// TIA Portal V18 export
FUNCTION "BYPASS DOS EQUIPAMENTOS" : Void   // FC12, LAD
{ S7_Optimized_Access := 'TRUE' }
// stored: SetENOAutomatically false
BEGIN

REGION Network 1: BYPASS GERAL E ESVAZIAMENTO DOS TRANSPORTADORES
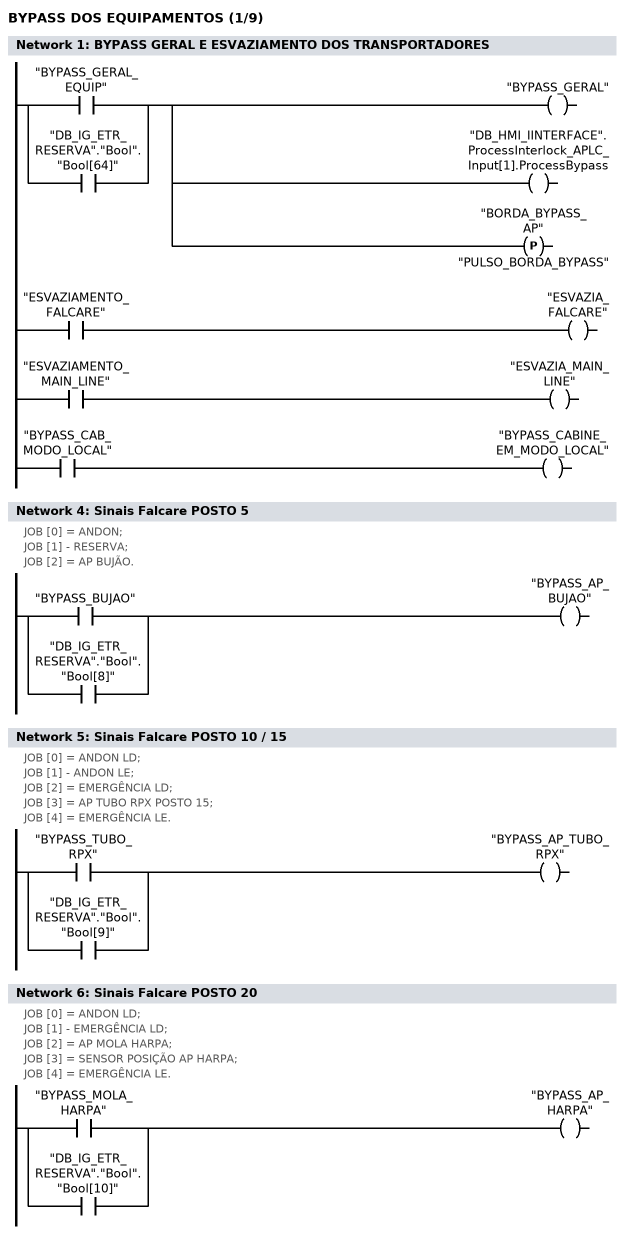
   "BYPASS_GERAL" := "BYPASS_GERAL_EQUIP" OR "DB_IG_ETR_RESERVA"."Bool"."Bool[64]";
   "DB_HMI_IINTERFACE".ProcessInterlock_APLC_Input[1].ProcessBypass := "BYPASS_GERAL";
   "BORDA_BYPASS_AP" := "BYPASS_GERAL" AND NOT "PULSO_BORDA_BYPASS";   // rising edge
   "PULSO_BORDA_BYPASS" := "BYPASS_GERAL";
   "ESVAZIA_FALCARE" := "ESVAZIAMENTO_FALCARE";
   "ESVAZIA_MAIN_LINE" := "ESVAZIAMENTO_MAIN_LINE";
   "BYPASS_CABINE_EM_MODO_LOCAL" := "BYPASS_CAB_MODO_LOCAL";
END_REGION

REGION Network 2: Sinais Falcare POSTO 1
   // JOB [0] = ANDON;
   // JOB [1] - EMERGÊNCIA;
END_REGION

REGION Network 3: Sinais Falcare VIVERK
   // JOB [0] = ANDON;
   // JOB [1] - EMERGÊNCIA;
END_REGION

REGION Network 4: Sinais Falcare POSTO 5
   // JOB [0] = ANDON;
   // JOB [1] - RESERVA;
   // JOB [2] = AP BUJÃO.
   RUNG wire#powerrail
      Contact( "BYPASS_BUJAO" )
      wire#w1
      Coil( "BYPASS_AP_BUJAO" )
   END_RUNG
   RUNG wire#powerrail
      Contact( "DB_IG_ETR_RESERVA"."Bool"."Bool[8]" )
   END_RUNG wire#w1
   // the same network as SCL:
   "BYPASS_AP_BUJAO" := "BYPASS_BUJAO" OR "DB_IG_ETR_RESERVA"."Bool"."Bool[8]";
END_REGION

REGION Network 5: Sinais Falcare POSTO 10 / 15
   // JOB [0] = ANDON LD;
   // JOB [1] - ANDON LE;
   // JOB [2] = EMERGÊNCIA LD;
   // JOB [3] = AP TUBO RPX POSTO 15;
   // JOB [4] = EMERGÊNCIA LE.
   RUNG wire#powerrail
      Contact( "BYPASS_TUBO_RPX" )
      wire#w1
      Coil( "BYPASS_AP_TUBO_RPX" )
   END_RUNG
   RUNG wire#powerrail
      Contact( "DB_IG_ETR_RESERVA"."Bool"."Bool[9]" )
   END_RUNG wire#w1
   // the same network as SCL:
   "BYPASS_AP_TUBO_RPX" := "BYPASS_TUBO_RPX" OR "DB_IG_ETR_RESERVA"."Bool"."Bool[9]";
END_REGION

REGION Network 6: Sinais Falcare POSTO 20
   // JOB [0] = ANDON LD;
   // JOB [1] - EMERGÊNCIA LD;
   // JOB [2] = AP MOLA HARPA;
   // JOB [3] = SENSOR POSIÇÃO AP HARPA;
   // JOB [4] = EMERGÊNCIA LE.
   RUNG wire#powerrail
      Contact( "BYPASS_MOLA_HARPA" )
      wire#w1
      Coil( "BYPASS_AP_HARPA" )
   END_RUNG
   RUNG wire#powerrail
      Contact( "DB_IG_ETR_RESERVA"."Bool"."Bool[10]" )
   END_RUNG wire#w1
   // the same network as SCL:
   "BYPASS_AP_HARPA" := "BYPASS_MOLA_HARPA" OR "DB_IG_ETR_RESERVA"."Bool"."Bool[10]";
END_REGION

REGION Network 7: Sinais Falcare POSTO 30
   // JOB [0] = ANDON LD;
   // JOB [1] = ANDON LE;
   // JOB [2] = EMERGENCIA;
   // JOB [3] = AP DA CARCAÇA;
   // JOB [4] = POSIÇÃO TALHA DIF.
   // JOB [5] = PY JUNTA.
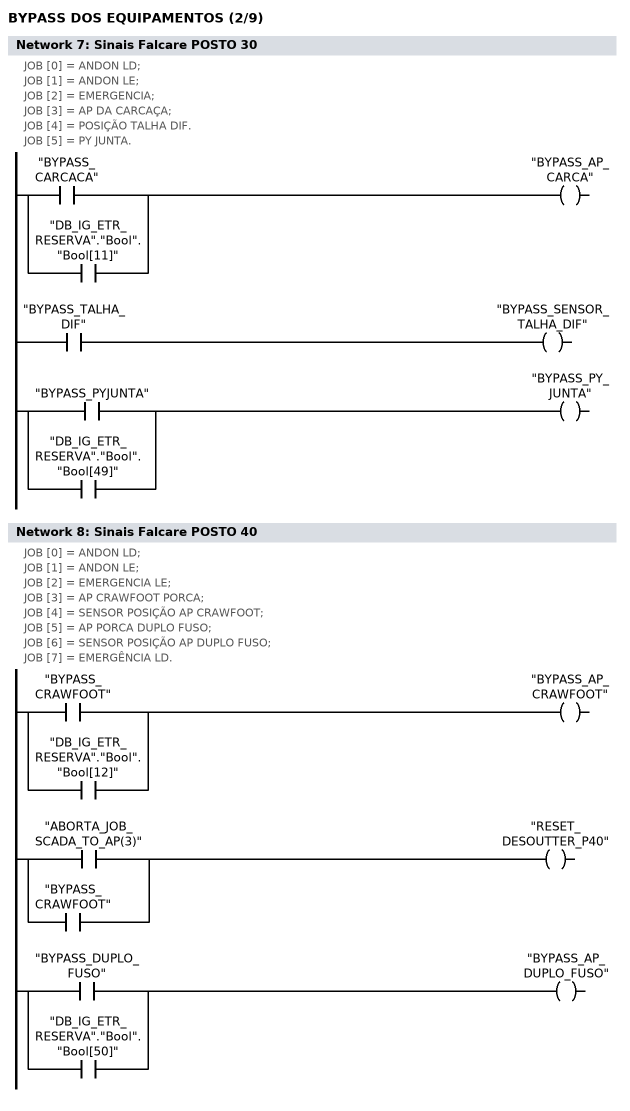
   RUNG wire#powerrail
      Contact( "BYPASS_CARCACA" )
      wire#w1
      Coil( "BYPASS_AP_CARCA" )
   END_RUNG
   RUNG wire#powerrail
      Contact( "DB_IG_ETR_RESERVA"."Bool"."Bool[11]" )
   END_RUNG wire#w1
   RUNG wire#powerrail
      Contact( "BYPASS_TALHA_DIF" )
      Coil( "BYPASS_SENSOR_TALHA_DIF" )
   END_RUNG
   RUNG wire#powerrail
      Contact( "BYPASS_PYJUNTA" )
      wire#w2
      Coil( "BYPASS_PY_JUNTA" )
   END_RUNG
   RUNG wire#powerrail
      Contact( "DB_IG_ETR_RESERVA"."Bool"."Bool[49]" )
   END_RUNG wire#w2
   // the same network as SCL:
   "BYPASS_AP_CARCA" := "BYPASS_CARCACA" OR "DB_IG_ETR_RESERVA"."Bool"."Bool[11]";
   "BYPASS_SENSOR_TALHA_DIF" := "BYPASS_TALHA_DIF";
   "BYPASS_PY_JUNTA" := "BYPASS_PYJUNTA" OR "DB_IG_ETR_RESERVA"."Bool"."Bool[49]";
END_REGION

REGION Network 8: Sinais Falcare POSTO 40
   // JOB [0] = ANDON LD;
   // JOB [1] = ANDON LE;
   // JOB [2] = EMERGENCIA LE;
   // JOB [3] = AP CRAWFOOT PORCA;
   // JOB [4] = SENSOR POSIÇÃO AP CRAWFOOT;
   // JOB [5] = AP PORCA DUPLO FUSO;
   // JOB [6] = SENSOR POSIÇÃO AP DUPLO FUSO;
   // JOB [7] = EMERGÊNCIA LD.
   RUNG wire#powerrail
      Contact( "BYPASS_CRAWFOOT" )
      wire#w1
      Coil( "BYPASS_AP_CRAWFOOT" )
   END_RUNG
   RUNG wire#powerrail
      Contact( "DB_IG_ETR_RESERVA"."Bool"."Bool[12]" )
   END_RUNG wire#w1
   RUNG wire#powerrail
      Contact( "ABORTA_JOB_SCADA_TO_AP(3)" )
      wire#w2
      Coil( "RESET_DESOUTTER_P40" )
   END_RUNG
   RUNG wire#powerrail
      Contact( "BYPASS_CRAWFOOT" )
   END_RUNG wire#w2
   RUNG wire#powerrail
      Contact( "BYPASS_DUPLO_FUSO" )
      wire#w3
      Coil( "BYPASS_AP_DUPLO_FUSO" )
   END_RUNG
   RUNG wire#powerrail
      Contact( "DB_IG_ETR_RESERVA"."Bool"."Bool[50]" )
   END_RUNG wire#w3
   // the same network as SCL:
   "BYPASS_AP_CRAWFOOT" := "BYPASS_CRAWFOOT" OR "DB_IG_ETR_RESERVA"."Bool"."Bool[12]";
   "RESET_DESOUTTER_P40" := "ABORTA_JOB_SCADA_TO_AP(3)" OR "BYPASS_CRAWFOOT";
   "BYPASS_AP_DUPLO_FUSO" := "BYPASS_DUPLO_FUSO" OR "DB_IG_ETR_RESERVA"."Bool"."Bool[50]";
END_REGION

REGION Network 9: Sinais Falcare POSTO 50 /55
   // JOB [0] = ANDON;
   // JOB [1] = EMERGENCIA;
   // JOB [2] = AP PORCA ESCONDIDA;
   // JOB [3] = SENSOR POSIÇÃO AP PORCA ESCONDIDA;
   // JOB [4] = AP PORCA SUPORTE DO CILINDRO;
   // JOB [5] = SENSOR POSIÇÃO AP SUPORTE DO CILINDRO;
   // JOB [6] = ANDON LD.
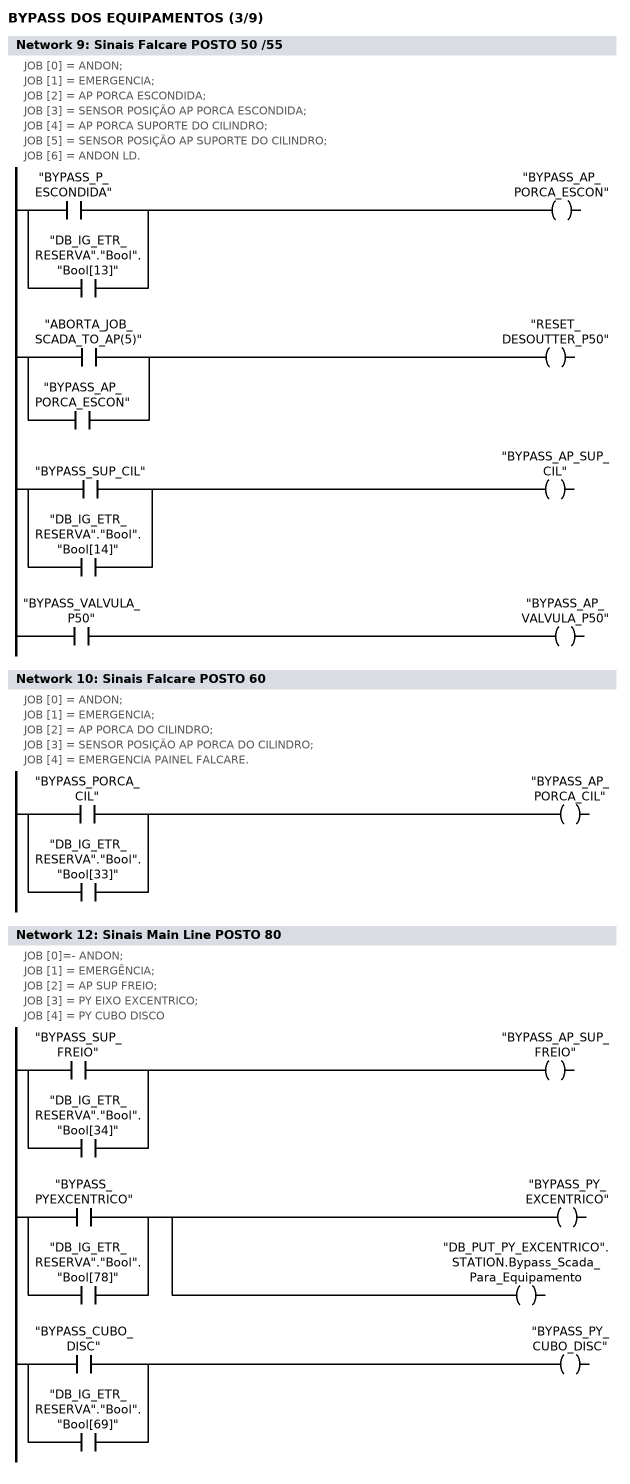
   RUNG wire#powerrail
      Contact( "BYPASS_P_ESCONDIDA" )
      wire#w1
      Coil( "BYPASS_AP_PORCA_ESCON" )
   END_RUNG
   RUNG wire#powerrail
      Contact( "DB_IG_ETR_RESERVA"."Bool"."Bool[13]" )
   END_RUNG wire#w1
   RUNG wire#powerrail
      Contact( "ABORTA_JOB_SCADA_TO_AP(5)" )
      wire#w2
      Coil( "RESET_DESOUTTER_P50" )
   END_RUNG
   RUNG wire#powerrail
      Contact( "BYPASS_AP_PORCA_ESCON" )
   END_RUNG wire#w2
   RUNG wire#powerrail
      Contact( "BYPASS_SUP_CIL" )
      wire#w3
      Coil( "BYPASS_AP_SUP_CIL" )
   END_RUNG
   RUNG wire#powerrail
      Contact( "DB_IG_ETR_RESERVA"."Bool"."Bool[14]" )
   END_RUNG wire#w3
   RUNG wire#powerrail
      Contact( "BYPASS_VALVULA_P50" )
      Coil( "BYPASS_AP_VALVULA_P50" )
   END_RUNG
   // the same network as SCL:
   "BYPASS_AP_PORCA_ESCON" := "BYPASS_P_ESCONDIDA" OR "DB_IG_ETR_RESERVA"."Bool"."Bool[13]";
   "RESET_DESOUTTER_P50" := "ABORTA_JOB_SCADA_TO_AP(5)" OR "BYPASS_AP_PORCA_ESCON";
   "BYPASS_AP_SUP_CIL" := "BYPASS_SUP_CIL" OR "DB_IG_ETR_RESERVA"."Bool"."Bool[14]";
   "BYPASS_AP_VALVULA_P50" := "BYPASS_VALVULA_P50";
END_REGION

REGION Network 10: Sinais Falcare POSTO 60
   // JOB [0] = ANDON;
   // JOB [1] = EMERGENCIA;
   // JOB [2] = AP PORCA DO CILINDRO;
   // JOB [3] = SENSOR POSIÇÃO AP PORCA DO CILINDRO;
   // JOB [4] = EMERGENCIA PAINEL FALCARE.
   RUNG wire#powerrail
      Contact( "BYPASS_PORCA_CIL" )
      wire#w1
      Coil( "BYPASS_AP_PORCA_CIL" )
   END_RUNG
   RUNG wire#powerrail
      Contact( "DB_IG_ETR_RESERVA"."Bool"."Bool[33]" )
   END_RUNG wire#w1
   // the same network as SCL:
   "BYPASS_AP_PORCA_CIL" := "BYPASS_PORCA_CIL" OR "DB_IG_ETR_RESERVA"."Bool"."Bool[33]";
END_REGION

REGION Network 11: Sinais Main Line POSTO 70 / 75
   // \\ JOB [0] - ANDON
END_REGION

REGION Network 12: Sinais Main Line POSTO 80
   // JOB [0]=- ANDON;
   // JOB [1] = EMERGÊNCIA;
   // JOB [2] = AP SUP FREIO;
   // JOB [3] = PY EIXO EXCENTRICO;
   // JOB [4] = PY CUBO DISCO
   RUNG wire#powerrail
      Contact( "BYPASS_SUP_FREIO" )
      wire#w1
      Coil( "BYPASS_AP_SUP_FREIO" )
   END_RUNG
   RUNG wire#powerrail
      Contact( "DB_IG_ETR_RESERVA"."Bool"."Bool[34]" )
   END_RUNG wire#w1
   RUNG wire#powerrail
      Contact( "BYPASS_PYEXCENTRICO" )
      wire#w2
      Coil( "BYPASS_PY_EXCENTRICO" )
   END_RUNG
   RUNG wire#powerrail
      Contact( "DB_IG_ETR_RESERVA"."Bool"."Bool[78]" )
   END_RUNG wire#w2
   RUNG wire#w2
      Coil( "DB_PUT_PY_EXCENTRICO".STATION.Bypass_Scada_Para_Equipamento )
   END_RUNG
   RUNG wire#powerrail
      Contact( "BYPASS_CUBO_DISC" )
      wire#w3
      Coil( "BYPASS_PY_CUBO_DISC" )
   END_RUNG
   RUNG wire#powerrail
      Contact( "DB_IG_ETR_RESERVA"."Bool"."Bool[69]" )
   END_RUNG wire#w3
   // the same network as SCL:
   "BYPASS_AP_SUP_FREIO" := "BYPASS_SUP_FREIO" OR "DB_IG_ETR_RESERVA"."Bool"."Bool[34]";
   "BYPASS_PY_EXCENTRICO" := "BYPASS_PYEXCENTRICO" OR "DB_IG_ETR_RESERVA"."Bool"."Bool[78]";
   "DB_PUT_PY_EXCENTRICO".STATION.Bypass_Scada_Para_Equipamento := "BYPASS_PY_EXCENTRICO";
   "BYPASS_PY_CUBO_DISC" := "BYPASS_CUBO_DISC" OR "DB_IG_ETR_RESERVA"."Bool"."Bool[69]";
END_REGION

REGION Network 13: Sinais Main Line POSTO 90 / 95
   // JOB [0] = ANDON;
   // JOB [1] = EMERGÊNCIA;
   // JOB [2] = AP HOLDER.
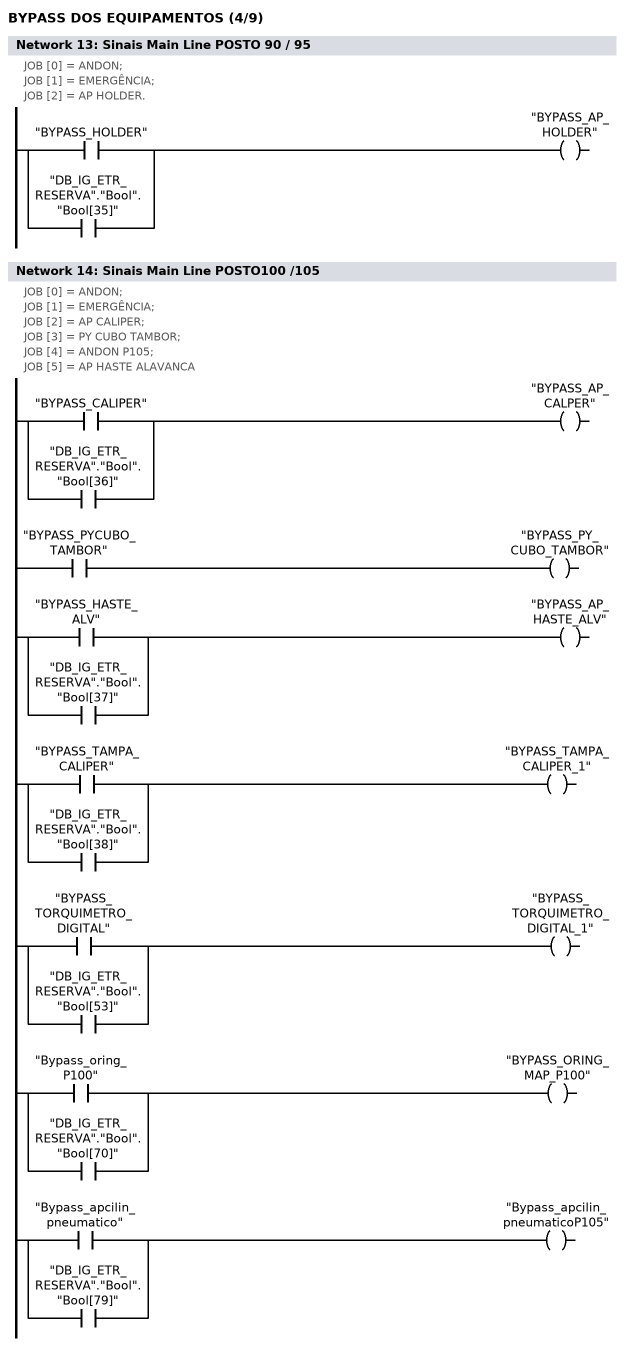
   RUNG wire#powerrail
      Contact( "BYPASS_HOLDER" )
      wire#w1
      Coil( "BYPASS_AP_HOLDER" )
   END_RUNG
   RUNG wire#powerrail
      Contact( "DB_IG_ETR_RESERVA"."Bool"."Bool[35]" )
   END_RUNG wire#w1
   // the same network as SCL:
   "BYPASS_AP_HOLDER" := "BYPASS_HOLDER" OR "DB_IG_ETR_RESERVA"."Bool"."Bool[35]";
END_REGION

REGION Network 14: Sinais Main Line POSTO100 /105
   // JOB [0] = ANDON;
   // JOB [1] = EMERGÊNCIA;
   // JOB [2] = AP CALIPER;
   // JOB [3] = PY CUBO TAMBOR;
   // JOB [4] = ANDON P105;
   // JOB [5] = AP HASTE ALAVANCA
   RUNG wire#powerrail
      Contact( "BYPASS_CALIPER" )
      wire#w1
      Coil( "BYPASS_AP_CALPER" )
   END_RUNG
   RUNG wire#powerrail
      Contact( "DB_IG_ETR_RESERVA"."Bool"."Bool[36]" )
   END_RUNG wire#w1
   RUNG wire#powerrail
      Contact( "BYPASS_PYCUBO_TAMBOR" )
      Coil( "BYPASS_PY_CUBO_TAMBOR" )
   END_RUNG
   RUNG wire#powerrail
      Contact( "BYPASS_HASTE_ALV" )
      wire#w2
      Coil( "BYPASS_AP_HASTE_ALV" )
   END_RUNG
   RUNG wire#powerrail
      Contact( "DB_IG_ETR_RESERVA"."Bool"."Bool[37]" )
   END_RUNG wire#w2
   RUNG wire#powerrail
      Contact( "BYPASS_TAMPA_CALIPER" )
      wire#w3
      Coil( "BYPASS_TAMPA_CALIPER_1" )
   END_RUNG
   RUNG wire#powerrail
      Contact( "DB_IG_ETR_RESERVA"."Bool"."Bool[38]" )
   END_RUNG wire#w3
   RUNG wire#powerrail
      Contact( "BYPASS_TORQUIMETRO_DIGITAL" )
      wire#w4
      Coil( "BYPASS_TORQUIMETRO_DIGITAL_1" )
   END_RUNG
   RUNG wire#powerrail
      Contact( "DB_IG_ETR_RESERVA"."Bool"."Bool[53]" )
   END_RUNG wire#w4
   RUNG wire#powerrail
      Contact( "Bypass_oring_P100" )
      wire#w5
      Coil( "BYPASS_ORING_MAP_P100" )
   END_RUNG
   RUNG wire#powerrail
      Contact( "DB_IG_ETR_RESERVA"."Bool"."Bool[70]" )
   END_RUNG wire#w5
   RUNG wire#powerrail
      Contact( "Bypass_apcilin_pneumatico" )
      wire#w6
      Coil( "Bypass_apcilin_pneumaticoP105" )
   END_RUNG
   RUNG wire#powerrail
      Contact( "DB_IG_ETR_RESERVA"."Bool"."Bool[79]" )
   END_RUNG wire#w6
   // the same network as SCL:
   "BYPASS_AP_CALPER" := "BYPASS_CALIPER" OR "DB_IG_ETR_RESERVA"."Bool"."Bool[36]";
   "BYPASS_PY_CUBO_TAMBOR" := "BYPASS_PYCUBO_TAMBOR";
   "BYPASS_AP_HASTE_ALV" := "BYPASS_HASTE_ALV" OR "DB_IG_ETR_RESERVA"."Bool"."Bool[37]";
   "BYPASS_TAMPA_CALIPER_1" := "BYPASS_TAMPA_CALIPER" OR "DB_IG_ETR_RESERVA"."Bool"."Bool[38]";
   "BYPASS_TORQUIMETRO_DIGITAL_1" := "BYPASS_TORQUIMETRO_DIGITAL" OR "DB_IG_ETR_RESERVA"."Bool"."Bool[53]";
   "BYPASS_ORING_MAP_P100" := "Bypass_oring_P100" OR "DB_IG_ETR_RESERVA"."Bool"."Bool[70]";
   "Bypass_apcilin_pneumaticoP105" := "Bypass_apcilin_pneumatico" OR "DB_IG_ETR_RESERVA"."Bool"."Bool[79]";
END_REGION

REGION Network 15: Sinais Main Line POSTO110 /115
   // JOB [0] = ANDON;
   // JOB [1] = SEG. BLOQUEIO CLP;
   // JOB [2] = AP CUBO;
   // JOB [3] = ANDON P115;
   // JOB [4] = CRAVADOR.
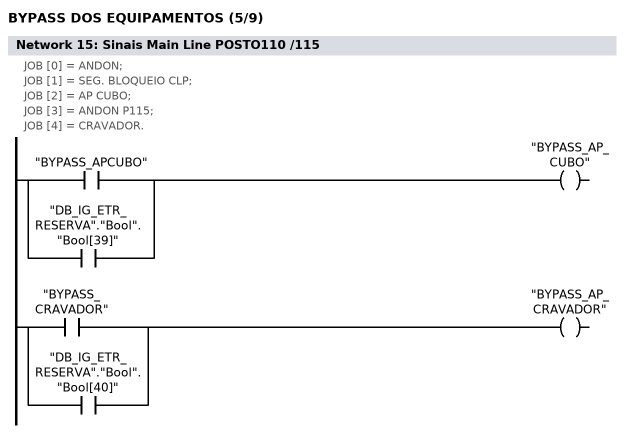
   RUNG wire#powerrail
      Contact( "BYPASS_APCUBO" )
      wire#w1
      Coil( "BYPASS_AP_CUBO" )
   END_RUNG
   RUNG wire#powerrail
      Contact( "DB_IG_ETR_RESERVA"."Bool"."Bool[39]" )
   END_RUNG wire#w1
   RUNG wire#powerrail
      Contact( "BYPASS_CRAVADOR" )
      wire#w2
      Coil( "BYPASS_AP_CRAVADOR" )
   END_RUNG
   RUNG wire#powerrail
      Contact( "DB_IG_ETR_RESERVA"."Bool"."Bool[40]" )
   END_RUNG wire#w2
   // the same network as SCL:
   "BYPASS_AP_CUBO" := "BYPASS_APCUBO" OR "DB_IG_ETR_RESERVA"."Bool"."Bool[39]";
   "BYPASS_AP_CRAVADOR" := "BYPASS_CRAVADOR" OR "DB_IG_ETR_RESERVA"."Bool"."Bool[40]";
END_REGION

REGION Network 16: Sinais Main Line POSTO120 /125
   // JOB [0] = ANDON;
   // JOB [1] - EMERGÊNCIA;
   // JOB [2] = AP INDICADOR;
   // JOB [3] = AP VALVULA;
   // JOB [4] = PY HELGE;
   // JOB [5] - ANDON P125;
   // JOB [6] - AP PORCA TERMINAL;
   // JOB [7] - AP FILTRO OLEO.
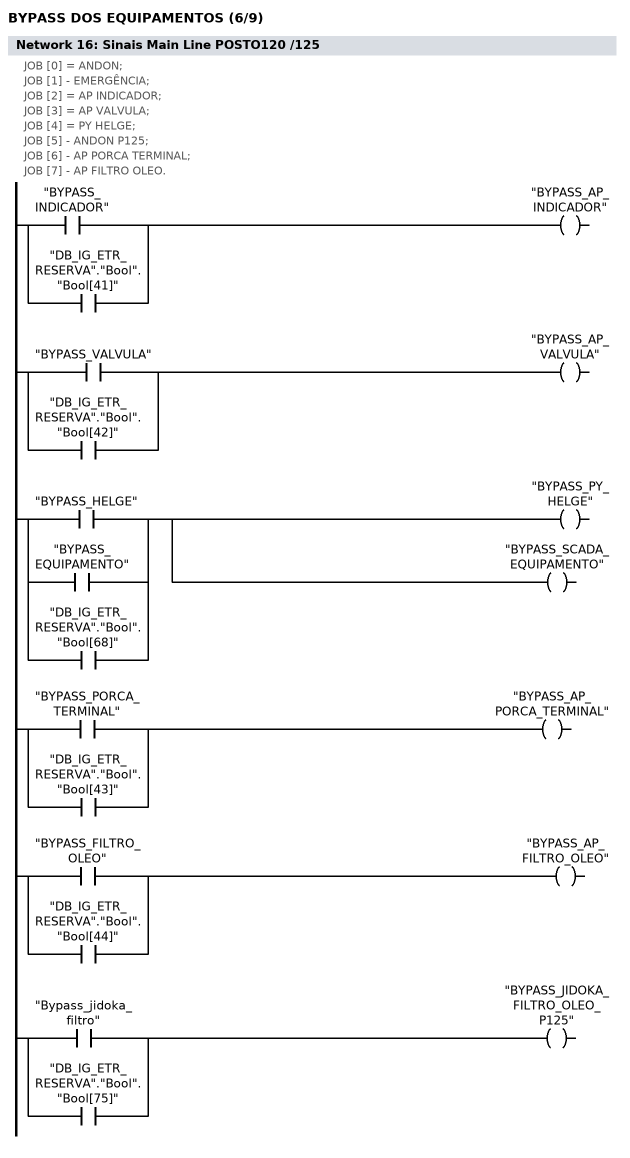
   RUNG wire#powerrail
      Contact( "BYPASS_INDICADOR" )
      wire#w1
      Coil( "BYPASS_AP_INDICADOR" )
   END_RUNG
   RUNG wire#powerrail
      Contact( "DB_IG_ETR_RESERVA"."Bool"."Bool[41]" )
   END_RUNG wire#w1
   RUNG wire#powerrail
      Contact( "BYPASS_VALVULA" )
      wire#w2
      Coil( "BYPASS_AP_VALVULA" )
   END_RUNG
   RUNG wire#powerrail
      Contact( "DB_IG_ETR_RESERVA"."Bool"."Bool[42]" )
   END_RUNG wire#w2
   RUNG wire#powerrail
      Contact( "BYPASS_HELGE" )
      wire#w3
      Coil( "BYPASS_PY_HELGE" )
   END_RUNG
   RUNG wire#powerrail
      Contact( "BYPASS_EQUIPAMENTO" )
   END_RUNG wire#w3
   RUNG wire#powerrail
      Contact( "DB_IG_ETR_RESERVA"."Bool"."Bool[68]" )
   END_RUNG wire#w3
   RUNG wire#w3
      Coil( "BYPASS_SCADA_EQUIPAMENTO" )
   END_RUNG
   RUNG wire#powerrail
      Contact( "BYPASS_PORCA_TERMINAL" )
      wire#w4
      Coil( "BYPASS_AP_PORCA_TERMINAL" )
   END_RUNG
   RUNG wire#powerrail
      Contact( "DB_IG_ETR_RESERVA"."Bool"."Bool[43]" )
   END_RUNG wire#w4
   RUNG wire#powerrail
      Contact( "BYPASS_FILTRO_OLEO" )
      wire#w5
      Coil( "BYPASS_AP_FILTRO_OLEO" )
   END_RUNG
   RUNG wire#powerrail
      Contact( "DB_IG_ETR_RESERVA"."Bool"."Bool[44]" )
   END_RUNG wire#w5
   RUNG wire#powerrail
      Contact( "Bypass_jidoka_filtro" )
      wire#w6
      Coil( "BYPASS_JIDOKA_FILTRO_OLEO_P125" )
   END_RUNG
   RUNG wire#powerrail
      Contact( "DB_IG_ETR_RESERVA"."Bool"."Bool[75]" )
   END_RUNG wire#w6
   // the same network as SCL:
   "BYPASS_AP_INDICADOR" := "BYPASS_INDICADOR" OR "DB_IG_ETR_RESERVA"."Bool"."Bool[41]";
   "BYPASS_AP_VALVULA" := "BYPASS_VALVULA" OR "DB_IG_ETR_RESERVA"."Bool"."Bool[42]";
   "BYPASS_PY_HELGE" := "BYPASS_HELGE" OR "BYPASS_EQUIPAMENTO" OR "DB_IG_ETR_RESERVA"."Bool"."Bool[68]";
   "BYPASS_SCADA_EQUIPAMENTO" := "BYPASS_PY_HELGE";
   "BYPASS_AP_PORCA_TERMINAL" := "BYPASS_PORCA_TERMINAL" OR "DB_IG_ETR_RESERVA"."Bool"."Bool[43]";
   "BYPASS_AP_FILTRO_OLEO" := "BYPASS_FILTRO_OLEO" OR "DB_IG_ETR_RESERVA"."Bool"."Bool[44]";
   "BYPASS_JIDOKA_FILTRO_OLEO_P125" := "Bypass_jidoka_filtro" OR "DB_IG_ETR_RESERVA"."Bool"."Bool[75]";
END_REGION

REGION Network 17: Sinais Main Line POSTO130
   // JOB [0] = ANDON;
   // JOB [1] = AP REDUÇÃO;
   // JOB [2] - AP FALNGE
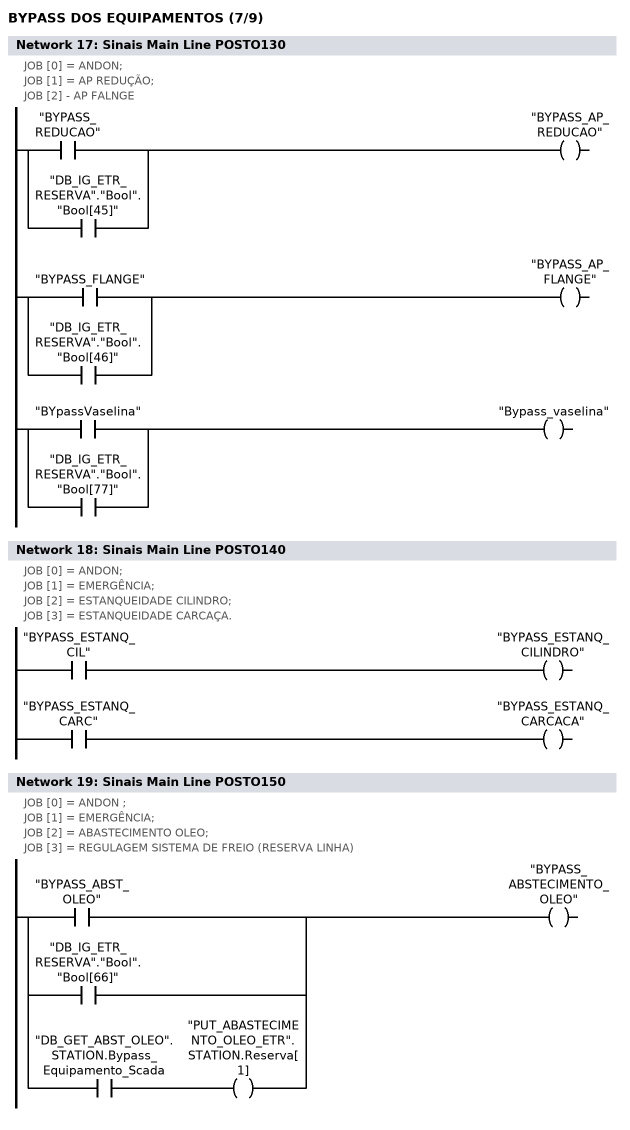
   RUNG wire#powerrail
      Contact( "BYPASS_REDUCAO" )
      wire#w1
      Coil( "BYPASS_AP_REDUCAO" )
   END_RUNG
   RUNG wire#powerrail
      Contact( "DB_IG_ETR_RESERVA"."Bool"."Bool[45]" )
   END_RUNG wire#w1
   RUNG wire#powerrail
      Contact( "BYPASS_FLANGE" )
      wire#w2
      Coil( "BYPASS_AP_FLANGE" )
   END_RUNG
   RUNG wire#powerrail
      Contact( "DB_IG_ETR_RESERVA"."Bool"."Bool[46]" )
   END_RUNG wire#w2
   RUNG wire#powerrail
      Contact( "BYpassVaselina" )
      wire#w3
      Coil( "Bypass_vaselina" )
   END_RUNG
   RUNG wire#powerrail
      Contact( "DB_IG_ETR_RESERVA"."Bool"."Bool[77]" )
   END_RUNG wire#w3
   // the same network as SCL:
   "BYPASS_AP_REDUCAO" := "BYPASS_REDUCAO" OR "DB_IG_ETR_RESERVA"."Bool"."Bool[45]";
   "BYPASS_AP_FLANGE" := "BYPASS_FLANGE" OR "DB_IG_ETR_RESERVA"."Bool"."Bool[46]";
   "Bypass_vaselina" := "BYpassVaselina" OR "DB_IG_ETR_RESERVA"."Bool"."Bool[77]";
END_REGION

REGION Network 18: Sinais Main Line POSTO140
   // JOB [0] = ANDON;
   // JOB [1] = EMERGÊNCIA;
   // JOB [2] = ESTANQUEIDADE CILINDRO;
   // JOB [3] = ESTANQUEIDADE CARCAÇA.
   RUNG wire#powerrail
      Contact( "BYPASS_ESTANQ_CIL" )
      Coil( "BYPASS_ESTANQ_CILINDRO" )
   END_RUNG
   RUNG wire#powerrail
      Contact( "BYPASS_ESTANQ_CARC" )
      Coil( "BYPASS_ESTANQ_CARCACA" )
   END_RUNG
   // the same network as SCL:
   "BYPASS_ESTANQ_CILINDRO" := "BYPASS_ESTANQ_CIL";
   "BYPASS_ESTANQ_CARCACA" := "BYPASS_ESTANQ_CARC";
END_REGION

REGION Network 19: Sinais Main Line POSTO150
   // JOB [0] = ANDON ;
   // JOB [1] = EMERGÊNCIA;
   // JOB [2] = ABASTECIMENTO OLEO;
   // JOB [3] = REGULAGEM SISTEMA DE FREIO (RESERVA LINHA)
   RUNG wire#powerrail
      Contact( "BYPASS_ABST_OLEO" )
      wire#w1
      Coil( "BYPASS_ABSTECIMENTO_OLEO" )
   END_RUNG
   RUNG wire#powerrail
      Contact( "DB_IG_ETR_RESERVA"."Bool"."Bool[66]" )
   END_RUNG wire#w1
   RUNG wire#powerrail
      Contact( "DB_GET_ABST_OLEO".STATION.Bypass_Equipamento_Scada )
      Coil( "PUT_ABASTECIMENTO_OLEO_ETR".STATION.Reserva[1] )
   END_RUNG wire#w1
   // the same network as SCL:
   "PUT_ABASTECIMENTO_OLEO_ETR".STATION.Reserva[1] := "DB_GET_ABST_OLEO".STATION.Bypass_Equipamento_Scada;
   "BYPASS_ABSTECIMENTO_OLEO" := "BYPASS_ABST_OLEO" OR "DB_IG_ETR_RESERVA"."Bool"."Bool[66]" OR "DB_GET_ABST_OLEO".STATION.Bypass_Equipamento_Scada;
END_REGION

REGION Network 20: Sinais Main Line Q.G
   // JOB [0] = ANDON;
   // JOB [1] = EMERGÊNCIA;
   // JOB [2] - EIXO PENDURADO;
   // JOB [3] - GAP PRESENTE CAB;
   // JOB [4] - GAP PRESENTE TAKT
END_REGION

REGION Network 21: Sinais Main Line EXPEDIÇÃO
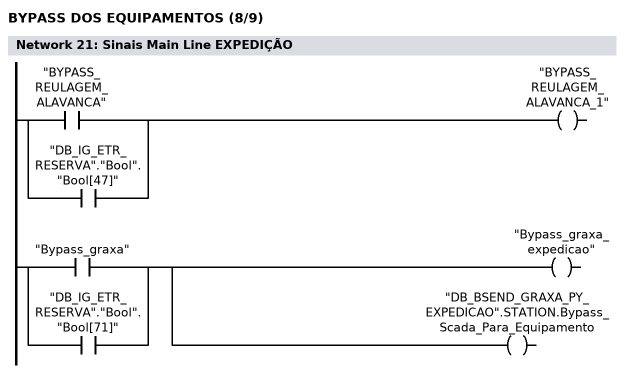
   RUNG wire#powerrail
      Contact( "BYPASS_REULAGEM_ALAVANCA" )
      wire#w1
      Coil( "BYPASS_REULAGEM_ALAVANCA_1" )
   END_RUNG
   RUNG wire#powerrail
      Contact( "DB_IG_ETR_RESERVA"."Bool"."Bool[47]" )
   END_RUNG wire#w1
   RUNG wire#powerrail
      Contact( "Bypass_graxa" )
      wire#w2
      Coil( "Bypass_graxa_expedicao" )
   END_RUNG
   RUNG wire#powerrail
      Contact( "DB_IG_ETR_RESERVA"."Bool"."Bool[71]" )
   END_RUNG wire#w2
   RUNG wire#w2
      Coil( "DB_BSEND_GRAXA_PY_EXPEDICAO".STATION.Bypass_Scada_Para_Equipamento )
   END_RUNG
   // the same network as SCL:
   "BYPASS_REULAGEM_ALAVANCA_1" := "BYPASS_REULAGEM_ALAVANCA" OR "DB_IG_ETR_RESERVA"."Bool"."Bool[47]";
   "Bypass_graxa_expedicao" := "Bypass_graxa" OR "DB_IG_ETR_RESERVA"."Bool"."Bool[71]";
   "DB_BSEND_GRAXA_PY_EXPEDICAO".STATION.Bypass_Scada_Para_Equipamento := "Bypass_graxa_expedicao";
END_REGION

REGION Network 22: BYPASS STATIONS
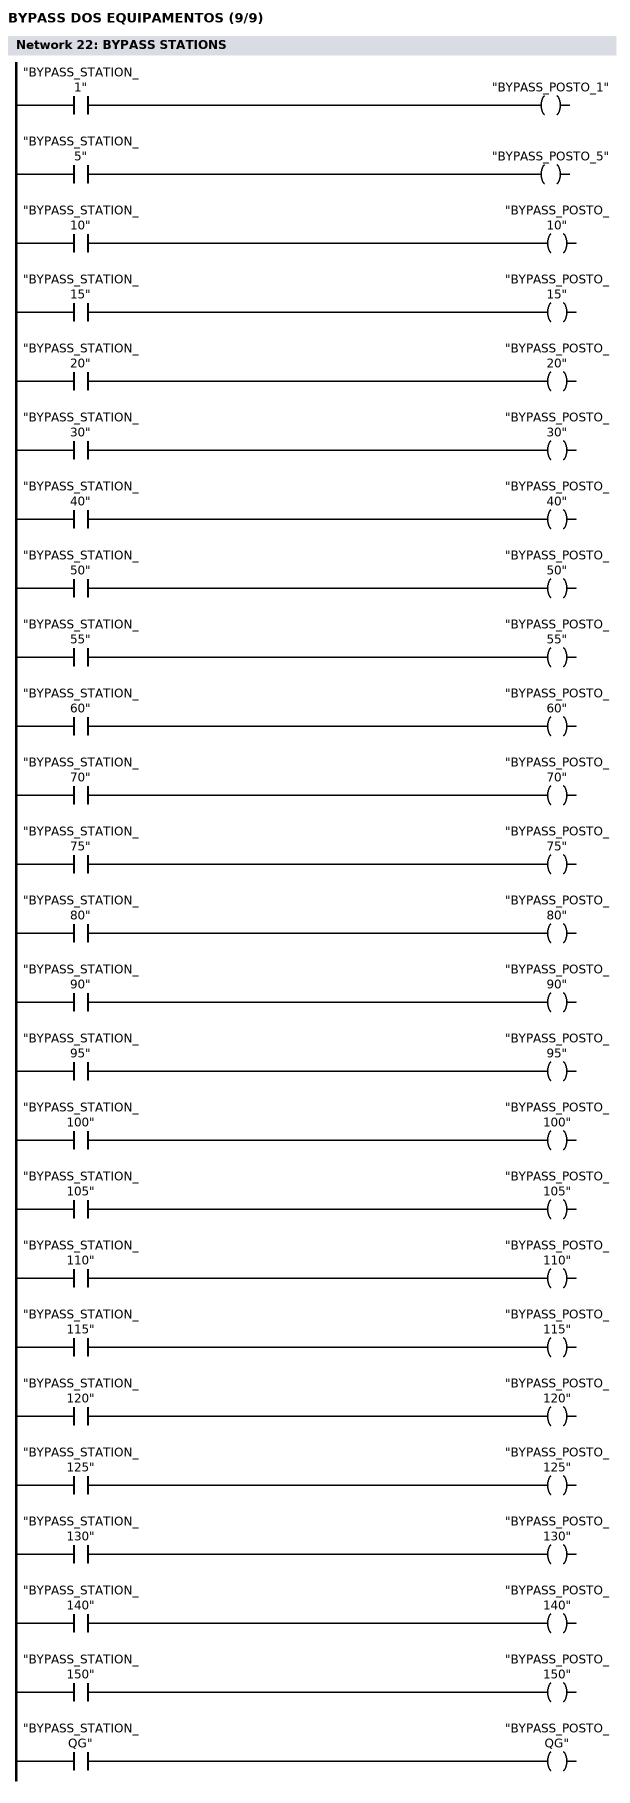
   RUNG wire#powerrail
      Contact( "BYPASS_STATION_1" )
      Coil( "BYPASS_POSTO_1" )
   END_RUNG
   RUNG wire#powerrail
      Contact( "BYPASS_STATION_5" )
      Coil( "BYPASS_POSTO_5" )
   END_RUNG
   RUNG wire#powerrail
      Contact( "BYPASS_STATION_10" )
      Coil( "BYPASS_POSTO_10" )
   END_RUNG
   RUNG wire#powerrail
      Contact( "BYPASS_STATION_15" )
      Coil( "BYPASS_POSTO_15" )
   END_RUNG
   RUNG wire#powerrail
      Contact( "BYPASS_STATION_20" )
      Coil( "BYPASS_POSTO_20" )
   END_RUNG
   RUNG wire#powerrail
      Contact( "BYPASS_STATION_30" )
      Coil( "BYPASS_POSTO_30" )
   END_RUNG
   RUNG wire#powerrail
      Contact( "BYPASS_STATION_40" )
      Coil( "BYPASS_POSTO_40" )
   END_RUNG
   RUNG wire#powerrail
      Contact( "BYPASS_STATION_50" )
      Coil( "BYPASS_POSTO_50" )
   END_RUNG
   RUNG wire#powerrail
      Contact( "BYPASS_STATION_55" )
      Coil( "BYPASS_POSTO_55" )
   END_RUNG
   RUNG wire#powerrail
      Contact( "BYPASS_STATION_60" )
      Coil( "BYPASS_POSTO_60" )
   END_RUNG
   RUNG wire#powerrail
      Contact( "BYPASS_STATION_70" )
      Coil( "BYPASS_POSTO_70" )
   END_RUNG
   RUNG wire#powerrail
      Contact( "BYPASS_STATION_75" )
      Coil( "BYPASS_POSTO_75" )
   END_RUNG
   RUNG wire#powerrail
      Contact( "BYPASS_STATION_80" )
      Coil( "BYPASS_POSTO_80" )
   END_RUNG
   RUNG wire#powerrail
      Contact( "BYPASS_STATION_90" )
      Coil( "BYPASS_POSTO_90" )
   END_RUNG
   RUNG wire#powerrail
      Contact( "BYPASS_STATION_95" )
      Coil( "BYPASS_POSTO_95" )
   END_RUNG
   RUNG wire#powerrail
      Contact( "BYPASS_STATION_100" )
      Coil( "BYPASS_POSTO_100" )
   END_RUNG
   RUNG wire#powerrail
      Contact( "BYPASS_STATION_105" )
      Coil( "BYPASS_POSTO_105" )
   END_RUNG
   RUNG wire#powerrail
      Contact( "BYPASS_STATION_110" )
      Coil( "BYPASS_POSTO_110" )
   END_RUNG
   RUNG wire#powerrail
      Contact( "BYPASS_STATION_115" )
      Coil( "BYPASS_POSTO_115" )
   END_RUNG
   RUNG wire#powerrail
      Contact( "BYPASS_STATION_120" )
      Coil( "BYPASS_POSTO_120" )
   END_RUNG
   RUNG wire#powerrail
      Contact( "BYPASS_STATION_125" )
      Coil( "BYPASS_POSTO_125" )
   END_RUNG
   RUNG wire#powerrail
      Contact( "BYPASS_STATION_130" )
      Coil( "BYPASS_POSTO_130" )
   END_RUNG
   RUNG wire#powerrail
      Contact( "BYPASS_STATION_140" )
      Coil( "BYPASS_POSTO_140" )
   END_RUNG
   RUNG wire#powerrail
      Contact( "BYPASS_STATION_150" )
      Coil( "BYPASS_POSTO_150" )
   END_RUNG
   RUNG wire#powerrail
      Contact( "BYPASS_STATION_QG" )
      Coil( "BYPASS_POSTO_QG" )
   END_RUNG
   // the same network as SCL:
   "BYPASS_POSTO_1" := "BYPASS_STATION_1";
   "BYPASS_POSTO_5" := "BYPASS_STATION_5";
   "BYPASS_POSTO_10" := "BYPASS_STATION_10";
   "BYPASS_POSTO_15" := "BYPASS_STATION_15";
   "BYPASS_POSTO_20" := "BYPASS_STATION_20";
   "BYPASS_POSTO_30" := "BYPASS_STATION_30";
   "BYPASS_POSTO_40" := "BYPASS_STATION_40";
   "BYPASS_POSTO_50" := "BYPASS_STATION_50";
   "BYPASS_POSTO_55" := "BYPASS_STATION_55";
   "BYPASS_POSTO_60" := "BYPASS_STATION_60";
   "BYPASS_POSTO_70" := "BYPASS_STATION_70";
   "BYPASS_POSTO_75" := "BYPASS_STATION_75";
   "BYPASS_POSTO_80" := "BYPASS_STATION_80";
   "BYPASS_POSTO_90" := "BYPASS_STATION_90";
   "BYPASS_POSTO_95" := "BYPASS_STATION_95";
   "BYPASS_POSTO_100" := "BYPASS_STATION_100";
   "BYPASS_POSTO_105" := "BYPASS_STATION_105";
   "BYPASS_POSTO_110" := "BYPASS_STATION_110";
   "BYPASS_POSTO_115" := "BYPASS_STATION_115";
   "BYPASS_POSTO_120" := "BYPASS_STATION_120";
   "BYPASS_POSTO_125" := "BYPASS_STATION_125";
   "BYPASS_POSTO_130" := "BYPASS_STATION_130";
   "BYPASS_POSTO_140" := "BYPASS_STATION_140";
   "BYPASS_POSTO_150" := "BYPASS_STATION_150";
   "BYPASS_POSTO_QG" := "BYPASS_STATION_QG";
END_REGION
END_FUNCTION
